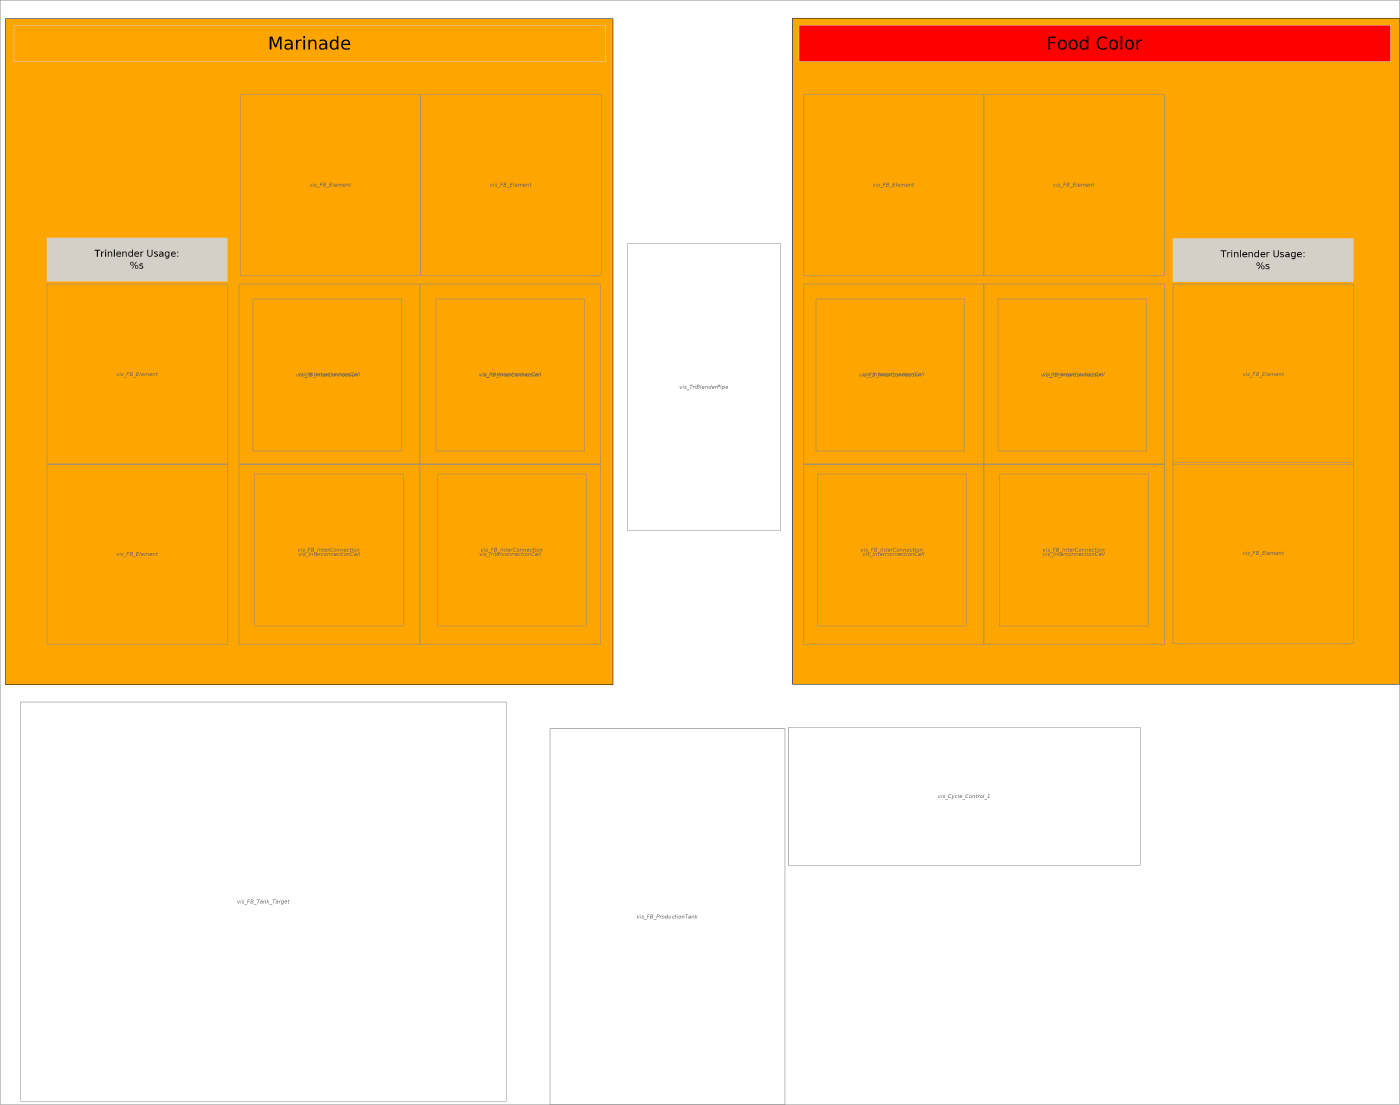
VISUALIZATION vis_Main  // 2638x2083
    Rectangle (1493,34 1145x1256)
    Frame (1513,178 341x341)
        shows vis_FB_Element(fb := fbElement[E_Element_List.eTank_3])
    Frame (1853,178 341x341)
        shows vis_FB_Element(fb := fbElement[E_Element_List.eTank_4])
    Frame (2210,535 341x341)
        shows vis_FB_Element(fb := fbElement[E_Element_List.eTriBlender_Color])
    Frame (2210,872 341x341)
        shows vis_FB_Element(fb := fbElement[E_Element_List.eLine_Color])
    Frame (1513,535 341x341)
        shows vis_InterconnectionCell()
    Frame (1853,535 341x341)
        shows vis_InterconnectionCell()
    Frame (1513,874 341x341)
        shows vis_InterconnectionCell()
    Frame (1853,874 341x341)
        shows vis_InterconnectionCell()
    Frame (1537,563 281x287)
        shows vis_FB_InterConnection(fb := fbIntCon_TriB_T3_Color)
    Frame (1880,563 281x287)
        shows vis_FB_InterConnection(fb := fbIntCon_TriB_T4_Color)
    Frame (1540,893 281x287)
        shows vis_FB_InterConnection(fb := fbIntCon_ProL_T3_Color)
    Frame (1883,893 281x287)
        shows vis_FB_InterConnection(fb := fbIntCon_ProL_T4_Color)
    Textfield (1505,47 1115x69), "Food Color"
    Group (10,35 1145x1256)
        Rectangle (0,0 1145x1256)
        Frame (442,143 341x341)
            shows vis_FB_Element(fb := fbElement[E_Element_List.eTank_1])
        Frame (782,143 341x341)
            shows vis_FB_Element(fb := fbElement[E_Element_List.eTank_2])
        Frame (78,500 341x341)
            shows vis_FB_Element(fb := fbElement[E_Element_List.eTriBlender_Marinada])
        Frame (78,839 341x341)
            shows vis_FB_Element(fb := fbElement[E_Element_List.eLine_Marinada])
        Frame (440,500 341x341)
            shows vis_InterconnectionCell()
        Frame (781,500 341x341)
            shows vis_InterconnectionCell()
        Frame (440,839 341x341)
            shows vis_InterconnectionCell()
        Frame (781,839 341x341)
            shows vis_InterconnectionCell()
        Frame (466,528 281x287)
            shows vis_FB_InterConnection(fb := fbIntCon_TriB_T1_Marin)
        Frame (811,528 281x287)
            shows vis_FB_InterConnection(fb := fbIntCon_TriB_T2_Marin)
        Frame (469,858 281x287)
            shows vis_FB_InterConnection(fb := fbIntCon_ProL_T1_Marin)
        Frame (814,858 281x287)
            shows vis_FB_InterConnection(fb := fbIntCon_ProL_T2_Marin)
        Textfield (16,12 1115x69), "Marinade"
        Textfield (78,413 340x82), "Trinlender Usage: %s", colour toggle: eTriBlenderUsage=E_TriBlenderUsage.eColor_Standby OR eTriBlenderUsage=E_TriBlenderUsage.eColor_T3 OR eTriBlenderUsage=E_TriBlenderUsage.eColor_T4, text list: 'TextList_TriBlenderUsage', text index: eTriBlenderUsage
    Textfield (2210,449 340x82), "Trinlender Usage: %s", colour toggle: eTriBlenderUsage=E_TriBlenderUsage.eMarinada_Standby OR eTriBlenderUsage=E_TriBlenderUsage.eMarinada_T1 OR eTriBlenderUsage=E_TriBlenderUsage.eMarinada_T2, text list: 'TextList_TriBlenderUsage', text index: eTriBlenderUsage
    Frame (1182,459 289x541)
        shows vis_TriBlenderPipe()
    Frame (1485,1371 664x260)
        shows vis_Cycle_Control_1(fb := fbTank1, sName := 'T1 Marinade')
    Frame (1036,1373 443x710)
        shows vis_FB_ProductionTank(fb := fbTank1)
    Frame (38,1323 916x753)
        shows vis_FB_Tank_Target(fb := fbTank1.fbTarget)
END_VISUALIZATION

(* stored: Version 1.1.0.1, ProductVersion 3.1.4024.12
   Visu vis_Main: Id {6e37a4b3-8f2f-410e-badf-675a7ad171d7} *)
